// TIA Portal V21 export
// export: Created 2026-08-21T20:18:54.114371Z, ExportSetting None, DisplayName Totally Integrated Automation Portal, DisplayVersion V21, DisplayName STEP 7 Professional, DisplayVersion V21, DisplayName STEP 7 Safety, DisplayVersion V21, DisplayName Tech WebApplication, DisplayVersion V21, DisplayName WinCC Basic/Comfort/Advanced, DisplayVersion V21, DisplayName WinCC Professional, DisplayVersion V21, DisplayName WinCC Unified, DisplayVersion V21
TYPE "typeMTPModuleTypePackageRevision"
TITLE = MTP-Versionierung / MTP versioning
// MTP Versionsinformation / MTP version information
   STRUCT
      ModuleTypePackageRevision { ExternalAccessible := 'False'; ExternalVisible := 'False'; ExternalWritable := 'False'} : String := '0.0.1';   // ModuleTypePackageRevision; Schema: Major.Minor.Patch / ModuleTypePackageRevision; scheme: Major.Minor.Patch
   END_STRUCT;
END_TYPE
